Fanuc KAREL source: KT00731.KL

PROGRAM KT00731
%NOLOCKGROUP
VAR
  ARG: ARRAY[4] OF INTEGER
  OUT: INTEGER
BEGIN
  OUT = ARRAY_LEN(ARG)
END KT00731
